Fanuc KAREL source: KT00774.KL

PROGRAM KT00774
%NOLOCKGROUP
VAR
  R1: REAL
  R2: REAL
  OUT: INTEGER
BEGIN
  R1 = 2.0
  R2 = 3.0
  R1 = 2.0
  R2 = 3.0
  OUT = ASIN(R1)
END KT00774
